(* CODESYS project visu_main_v0.export

Project tree, tasks and I/O mapping:
  visualisation Visu_Main
*)

// /Visu_Main
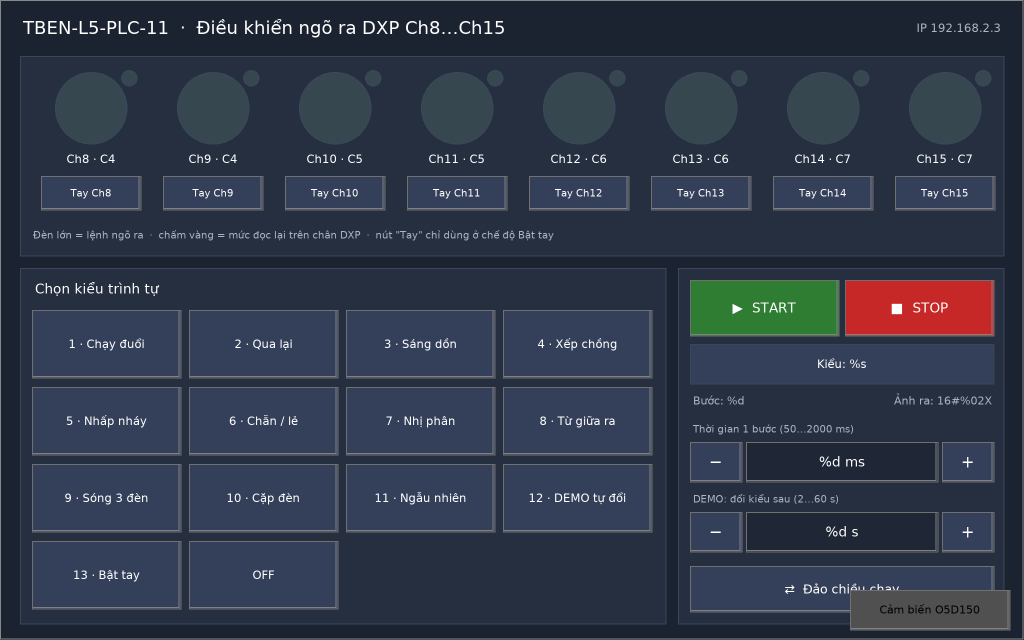
VISUALIZATION Visu_Main  // 1024x640
    Rectangle (0,0 1024x640)
    Rectangle (20,8 760x40), "TBEN-L5-PLC-11 · Điều khiển ngõ ra DXP Ch8…Ch15"
    Rectangle (784,8 220x40), "IP 192.168.2.3"
    RoundedRectangle (20,56 984x200)
    Ellipse (55,72 72x72), colour toggle: GVL_HMI.axOut[0]
    Ellipse (121,70 16x16), colour toggle: GVL_HMI.axFb[0]
    Rectangle (37,148 108x22), "Ch8 · C4"
    Button (41,176 100x34), "Tay Ch8", colour toggle: GVL_HMI.axManual[0], input disabled if: GVL_HMI.xNotManual
        toggle GVL_HMI.axManual[0]
    Ellipse (177,72 72x72), colour toggle: GVL_HMI.axOut[1]
    Ellipse (243,70 16x16), colour toggle: GVL_HMI.axFb[1]
    Rectangle (159,148 108x22), "Ch9 · C4"
    Button (163,176 100x34), "Tay Ch9", colour toggle: GVL_HMI.axManual[1], input disabled if: GVL_HMI.xNotManual
        toggle GVL_HMI.axManual[1]
    Ellipse (299,72 72x72), colour toggle: GVL_HMI.axOut[2]
    Ellipse (365,70 16x16), colour toggle: GVL_HMI.axFb[2]
    Rectangle (281,148 108x22), "Ch10 · C5"
    Button (285,176 100x34), "Tay Ch10", colour toggle: GVL_HMI.axManual[2], input disabled if: GVL_HMI.xNotManual
        toggle GVL_HMI.axManual[2]
    Ellipse (421,72 72x72), colour toggle: GVL_HMI.axOut[3]
    Ellipse (487,70 16x16), colour toggle: GVL_HMI.axFb[3]
    Rectangle (403,148 108x22), "Ch11 · C5"
    Button (407,176 100x34), "Tay Ch11", colour toggle: GVL_HMI.axManual[3], input disabled if: GVL_HMI.xNotManual
        toggle GVL_HMI.axManual[3]
    Ellipse (543,72 72x72), colour toggle: GVL_HMI.axOut[4]
    Ellipse (609,70 16x16), colour toggle: GVL_HMI.axFb[4]
    Rectangle (525,148 108x22), "Ch12 · C6"
    Button (529,176 100x34), "Tay Ch12", colour toggle: GVL_HMI.axManual[4], input disabled if: GVL_HMI.xNotManual
        toggle GVL_HMI.axManual[4]
    Ellipse (665,72 72x72), colour toggle: GVL_HMI.axOut[5]
    Ellipse (731,70 16x16), colour toggle: GVL_HMI.axFb[5]
    Rectangle (647,148 108x22), "Ch13 · C6"
    Button (651,176 100x34), "Tay Ch13", colour toggle: GVL_HMI.axManual[5], input disabled if: GVL_HMI.xNotManual
        toggle GVL_HMI.axManual[5]
    Ellipse (787,72 72x72), colour toggle: GVL_HMI.axOut[6]
    Ellipse (853,70 16x16), colour toggle: GVL_HMI.axFb[6]
    Rectangle (769,148 108x22), "Ch14 · C7"
    Button (773,176 100x34), "Tay Ch14", colour toggle: GVL_HMI.axManual[6], input disabled if: GVL_HMI.xNotManual
        toggle GVL_HMI.axManual[6]
    Ellipse (909,72 72x72), colour toggle: GVL_HMI.axOut[7]
    Ellipse (975,70 16x16), colour toggle: GVL_HMI.axFb[7]
    Rectangle (891,148 108x22), "Ch15 · C7"
    Button (895,176 100x34), "Tay Ch15", colour toggle: GVL_HMI.axManual[7], input disabled if: GVL_HMI.xNotManual
        toggle GVL_HMI.axManual[7]
    Rectangle (30,222 960x26), "Đèn lớn = lệnh ngõ ra · chấm vàng = mức đọc lại trên chân DXP · nút "Tay" chỉ dùng ở chế độ Bật tay"
    RoundedRectangle (20,268 646x356)
    Rectangle (32,274 600x30), "Chọn kiểu trình tự"
    Button (32,310 149x68), "1 · Chạy đuổi", colour toggle: GVL_HMI.axModeSel[1]
        OnMouseClick: execute { GVL_HMI.iModeSel := 1; }
    Button (189,310 149x68), "2 · Qua lại", colour toggle: GVL_HMI.axModeSel[2]
        OnMouseClick: execute { GVL_HMI.iModeSel := 2; }
    Button (346,310 149x68), "3 · Sáng dồn", colour toggle: GVL_HMI.axModeSel[3]
        OnMouseClick: execute { GVL_HMI.iModeSel := 3; }
    Button (503,310 149x68), "4 · Xếp chồng", colour toggle: GVL_HMI.axModeSel[4]
        OnMouseClick: execute { GVL_HMI.iModeSel := 4; }
    Button (32,387 149x68), "5 · Nhấp nháy", colour toggle: GVL_HMI.axModeSel[5]
        OnMouseClick: execute { GVL_HMI.iModeSel := 5; }
    Button (189,387 149x68), "6 · Chẵn / lẻ", colour toggle: GVL_HMI.axModeSel[6]
        OnMouseClick: execute { GVL_HMI.iModeSel := 6; }
    Button (346,387 149x68), "7 · Nhị phân", colour toggle: GVL_HMI.axModeSel[7]
        OnMouseClick: execute { GVL_HMI.iModeSel := 7; }
    Button (503,387 149x68), "8 · Từ giữa ra", colour toggle: GVL_HMI.axModeSel[8]
        OnMouseClick: execute { GVL_HMI.iModeSel := 8; }
    Button (32,464 149x68), "9 · Sóng 3 đèn", colour toggle: GVL_HMI.axModeSel[9]
        OnMouseClick: execute { GVL_HMI.iModeSel := 9; }
    Button (189,464 149x68), "10 · Cặp đèn", colour toggle: GVL_HMI.axModeSel[10]
        OnMouseClick: execute { GVL_HMI.iModeSel := 10; }
    Button (346,464 149x68), "11 · Ngẫu nhiên", colour toggle: GVL_HMI.axModeSel[11]
        OnMouseClick: execute { GVL_HMI.iModeSel := 11; }
    Button (503,464 149x68), "12 · DEMO tự đổi", colour toggle: GVL_HMI.axModeSel[12]
        OnMouseClick: execute { GVL_HMI.iModeSel := 12; }
    Button (32,541 149x68), "13 · Bật tay", colour toggle: GVL_HMI.axModeSel[13]
        OnMouseClick: execute { GVL_HMI.iModeSel := 13; }
    Button (189,541 149x68), "OFF", colour toggle: GVL_HMI.axModeSel[0]
        OnMouseClick: execute { GVL_HMI.iModeSel := 0; }
    RoundedRectangle (678,268 326x356)
    Button (690,280 149x56), "▶ START"
        OnMouseClick: execute { GVL_HMI.xCmdStart := TRUE; }
    Button (845,280 149x56), "■ STOP"
        OnMouseClick: execute { GVL_HMI.xCmdStop := TRUE; }
    RoundedRectangle (690,344 304x40), "Kiểu: %s", text variable: GVL_HMI.sModeName, colour toggle: GVL_HMI.xRunning
    Rectangle (690,388 150x26), "Bước: %d", text variable: GVL_HMI.uiStep
    Rectangle (845,388 150x26), "Ảnh ra: 16#%02X", text variable: GVL_HMI.byOut
    Rectangle (690,418 304x22), "Thời gian 1 bước (50…2000 ms)"
    Button (690,442 52x40), "−"
        OnMouseClick: execute { GVL_HMI.udiStepMs := GVL_HMI.udiStepMs - MIN(GVL_HMI.udiStepMs, 50); }
    Button (746,442 192x40), "%d ms", text variable: GVL_HMI.udiStepMs
        OnMouseClick: write GVL_HMI.udiStepMs via VisuDialogs.Numpad, min 50, max 2000, title "Thời gian bước [ms]"
    Button (942,442 52x40), "+"
        OnMouseClick: execute { GVL_HMI.udiStepMs := GVL_HMI.udiStepMs + 50; }
    Rectangle (690,488 304x22), "DEMO: đổi kiểu sau (2…60 s)"
    Button (690,512 52x40), "−"
        OnMouseClick: execute { GVL_HMI.udiDemoS := GVL_HMI.udiDemoS - MIN(GVL_HMI.udiDemoS, 1); }
    Button (746,512 192x40), "%d s", text variable: GVL_HMI.udiDemoS
        OnMouseClick: write GVL_HMI.udiDemoS via VisuDialogs.Numpad, min 2, max 60, title "Thời gian giữ mỗi kiểu [s]"
    Button (942,512 52x40), "+"
        OnMouseClick: execute { GVL_HMI.udiDemoS := GVL_HMI.udiDemoS + 1; }
    Button (690,566 304x46), "⇄ Đảo chiều chạy", colour toggle: GVL_HMI.xReverse
        toggle GVL_HMI.xReverse
    Button (850,590 160x40), "Cảm biến O5D150"
        OnMouseClick:  Assign=Visu_IOL_O5D150, Type=Assignment
END_VISUALIZATION
